(* IEC 61131-3 sources: Test-Git_ESME26/TestProgettoESME_26.fbsproj/PacDriveLib Migration/Motion/Homing/PDL_FB_Home.fb.st^, 21 files *)

(* ---- CallFb.meth.st ---- *)
{attribute 'conditionalshow_all_locals'}
METHOD PRIVATE CallFb
VAR_INPUT
END_VAR

CASE etHomeOpMode OF
	PDL_ET_HomeOpMode.TouchProbe:	(* HomeTP *)
		IF (stReducedVelocity_loc.i_xEnableReducedVelocity AND NOT stReducedVelocity_loc.i_xOnlyLimitCheck) THEN
			lrUsedVelocity := MIN(stReducedVelocity_loc.i_lrMaxReducedVelocity, stTouchProbe_loc.i_lrVel);
		ELSE
			lrUsedVelocity := stTouchProbe_loc.i_lrVel;
		END_IF
		fbHomeTP(	i_xEnable			:= xFbEnable,
					i_ifDrive			:= i_ifDrive,
					i_ifTouchProbe		:= stTouchProbe_loc.i_ifTouchProbe,
					i_etMode			:= etHomeTpMode,
					i_lrOffset			:= stTouchProbe_loc.i_lrOffset,
					i_lrMaxTravel		:= stTouchProbe_loc.i_lrMaxTravel,
					i_lrHomePosition	:= stTouchProbe_loc.i_lrHomePosition,
					i_lrVel				:= lrUsedVelocity,
					i_lrAcc				:= stTouchProbe_loc.i_lrAcc,
					i_lrDec				:= stTouchProbe_loc.i_lrDec,
					i_lrJerk			:= stTouchProbe_loc.i_lrJerk,
					i_xHwLimitNeg		:= i_xHwLimitNeg,
					i_xHwLimitPos		:= i_xHwLimitPos,
					i_xRotativeSystem	:= stTouchProbe_loc.i_xRotativeSystem,
					i_xStart			:= TRUE,
					q_xActive			=> xFbActive,
					q_xReady			=> ,
					q_etDiag			=> THIS^.etDiagBuffer,
					q_etDiagExt			=> ,
					q_sMsg				=> ,
					q_xMotionInstructionActive => ,
					q_lrPosition		=> ,
					q_xHomeOk			=> xFbHomeOk);
		THIS^.HomeTpDiagTranslation();

	PDL_ET_HomeOpMode.Sensor:	(* HomeIN *)
		IF (stReducedVelocity_loc.i_xEnableReducedVelocity AND NOT stReducedVelocity_loc.i_xOnlyLimitCheck) THEN
			lrUsedVelocity := MIN(stReducedVelocity_loc.i_lrMaxReducedVelocity, stSensor_loc.i_lrVel);
		ELSE
			lrUsedVelocity := stSensor_loc.i_lrVel;
		END_IF
		THIS^.fbHomeIn(	i_xEnable			:= xFbEnable,
					i_ifDrive			:= i_ifDrive,
					i_xSensor			:= stSensor_loc.i_xSensor,
					i_etMode			:= etHomeInMode,
					i_lrOffset			:= stSensor_loc.i_lrOffset,
					i_lrMaxTravel		:= stSensor_loc.i_lrMaxTravel,
					i_lrHomePosition	:= stSensor_loc.i_lrHomePosition,
					i_lrVel				:= lrUsedVelocity,
					i_lrAcc				:= stSensor_loc.i_lrAcc,
					i_lrDec				:= stSensor_loc.i_lrDec,
					i_lrJerk			:= stSensor_loc.i_lrJerk,
					i_xHwLimitNeg		:= i_xHwLimitNeg,
					i_xHwLimitPos		:= i_xHwLimitPos,
					i_xRotativeSystem	:= stSensor_loc.i_xRotativeSystem,
					i_xStart			:= xStartHomeIn,
					q_xActive			=> xFbActive,
					q_xReady			=> ,
					q_etDiag			=> THIS^.etDiagBuffer,
					q_etDiagExt			=> ,
					q_sMsg				=> ,
					q_xMotionInstructionActive => ,
					q_lrPosition		=> ,
					q_xHomeOk			=> xFbHomeOk);
		THIS^.HomeInDiagTranslation();

	PDL_ET_HomeOpMode.LimitSwitch:	(* HomeLS *)
		IF (stReducedVelocity_loc.i_xEnableReducedVelocity AND NOT stReducedVelocity_loc.i_xOnlyLimitCheck) THEN
			lrUsedVelocity := MIN(stReducedVelocity_loc.i_lrMaxReducedVelocity, stLimitSwitch_loc.i_lrVel);
		ELSE
			lrUsedVelocity := stLimitSwitch_loc.i_lrVel;
		END_IF
		IF (stLimitSwitch_loc.i_lrLowVel = 0.0) THEN
			lrLowVelocity := lrUsedVelocity;
		ELSE
			IF (stReducedVelocity_loc.i_xEnableReducedVelocity AND NOT stReducedVelocity_loc.i_xOnlyLimitCheck) THEN
				lrLowVelocity := MIN(stReducedVelocity_loc.i_lrMaxReducedVelocity, stLimitSwitch_loc.i_lrLowVel);
			ELSE
				lrLowVelocity := stLimitSwitch_loc.i_lrLowVel;
			END_IF
		END_IF
		fbHomeLS(	i_xEnable			:= xFbEnable,
					i_ifDrive			:= i_ifDrive,
					i_etMode			:= etHomeLimitSwitchMode,
					i_lrOffset			:= stLimitSwitch_loc.i_lrOffset,
					i_lrMaxTravel		:= stLimitSwitch_loc.i_lrMaxTravel,
					i_lrHomePosition	:= stLimitSwitch_loc.i_lrHomePosition,
					i_lrVel				:= lrUsedVelocity,
					i_lrLowVel			:= lrLowVelocity,
					i_lrAcc				:= stLimitSwitch_loc.i_lrAcc,
					i_lrDec				:= stLimitSwitch_loc.i_lrDec,
					i_lrJerk			:= stLimitSwitch_loc.i_lrJerk,
					i_xHwLimitNeg		:= i_xHwLimitNeg,
					i_xHwLimitPos		:= i_xHwLimitPos,
					i_xStart			:= TRUE,
					q_xActive			=> xFbActive,
					q_xReady			=> ,
					q_etDiag			=> THIS^.etDiagBuffer,
					q_etDiagExt			=> ,
					q_sMsg				=> ,
					q_xMotionInstructionActive => ,
					q_lrPosition		=> ,
					q_xHomeOk			=> xFbHomeOk);
		THIS^.HomeLSDiagTranslation();

	PDL_ET_HomeOpMode.Torque:	(* HomeTorque *)
		IF (stReducedVelocity_loc.i_xEnableReducedVelocity AND NOT stReducedVelocity_loc.i_xOnlyLimitCheck) THEN
			lrUsedVelocity := MIN(stReducedVelocity_loc.i_lrMaxReducedVelocity, stTorque_loc.i_lrVel);
		ELSE
			lrUsedVelocity := stTorque_loc.i_lrVel;
		END_IF
		fbHomeTorque(	i_xEnable			:= xFbEnable,
						i_ifDrive			:= i_ifDrive,
						i_lrMaxTorque		:= stTorque_loc.i_lrMaxTorque,
						i_diTorqueTime		:= stTorque_loc.i_diTorqueTime,
						i_lrLowLimit		:= -2147483648.0,
						i_lrHighLimit		:= 2147483648.0,
						i_etMode			:= etHomeTorqueMode,
						i_lrOffset			:= stTorque_loc.i_lrOffset,
						i_lrMaxTravel		:= stTorque_loc.i_lrMaxTravel,
						i_lrHomePosition	:= stTorque_loc.i_lrHomePosition,
						i_lrVel				:= lrUsedVelocity,
						i_lrAcc				:= stTorque_loc.i_lrAcc,
						i_lrDec				:= stTorque_loc.i_lrDec,
						i_lrJerk			:= stTorque_loc.i_lrJerk,
						i_xStart			:= TRUE,
						q_xActive			=> xFbActive,
						q_xReady			=> ,
						q_etDiag			=> THIS^.etDiagBuffer,
						q_etDiagExt			=> ,
						q_sMsg				=> ,
						q_xMotionInstructionActive => ,
						q_lrPosition		=> ,
						q_xHomeOk			=> xFbHomeOk);
		THIS^.HomeTorqueDiagTranslation();

	PDL_ET_HomeOpMode.Force:	(* HomeForce *)
			;

	PDL_ET_HomeOpMode.MoveOnPos:	(* Home to a Position *)
		IF (stReducedVelocity_loc.i_xEnableReducedVelocity AND NOT stReducedVelocity_loc.i_xOnlyLimitCheck) THEN
			lrUsedVelocity := MIN(stReducedVelocity_loc.i_lrMaxReducedVelocity, stMoveOnPos_loc.i_lrVel);
		ELSE
			lrUsedVelocity := stMoveOnPos_loc.i_lrVel;
		END_IF

		THIS^.fbVarioPosJerk(	i_xEnable			:= xFbEnable,
						i_ifDrive			:= i_ifDrive,
						i_xStart			:= fbVarioPosJerk.q_xActive AND TRUE,
						i_xStop				:= FALSE,
						i_lrTarget			:= lrPositionOpmMoveOnPos,
						i_lrVel				:= lrUsedVelocity,
						i_lrAcc				:= stMoveOnPos_loc.i_lrAcc,
						i_lrDec				:= stMoveOnPos_loc.i_lrDec,
						i_lrJerk			:= stMoveOnPos_loc.i_lrJerk,
						i_etPosMode			:= SEL(stMoveOnPos_loc.i_xRotativeSystem, PDL_ET_PosMode.Absolute, PDL_ET_PosMode.Relative),
						q_xActive			=> xFbActive,
						q_xReady			=> ,
						q_etDiag			=> THIS^.etDiagBuffer,
						q_etDiagExt			=> ,
						q_sMsg				=> ,
						q_xMotionInstructionActive => ,
						q_lrPosition		=> ,
						q_xInPosition		=> xFbHomeOk);

		THIS^.HomeMoveOnPosDiagTranslation();

		fbTrigStop(CLK:= xFbEnable AND (i_ifDrive.etAxisState = MOIN.ET_AxisState.Stopping));
		IF fbTrigStop.Q THEN
			xControllerStop :=  TRUE;
			xFbEnable := FALSE;
		END_IF

		// Clean up as soon as VarioPos is finished
		IF NOT xFbActive THEN
			// check, if VarioPos was aborted by MC_Stop OR MC_Halt
			IF xControllerStop THEN
				SetDiagOutput(	i_etDiag	:= GD.ET_Diag.HomingFailed,
								i_etDiagExt := PDL_ET_DiagExt.OutsideExecutionOfControllerStopSet,
								i_sMsg		:= 'MC_Stop OR MC_Halt was executed during homing active');
			ELSE
				IF stMoveOnPos_loc.i_lrPeriod > 0 AND stMoveOnPos_loc.i_xRotativeSystem THEN
					THIS^.fbSetPosIntern(
						Axis     := i_ifDrive,
						Position := stMoveOnPos_loc.i_lrTarget,
						Relative := FALSE,
						Execute  := TRUE);

					IF THIS^.fbSetPosIntern.Error THEN
							SetDiagOutput(	i_etDiag	:= GD.ET_Diag.UnexpectedProgramBehavior,
											i_etDiagExt := PDL_ET_DiagExt.UnexpectedFeedback,
											i_sMsg      := CONCAT('FB_Home error: MC_Setposition.ErrorID: ', PLCO.FC_EtResultToString(THIS^.fbSetPosIntern.ErrorID)));
					END_IF
					THIS^.fbSetPosIntern(Execute  := FALSE);
				END_IF
			END_IF
		END_IF

	PDL_ET_HomeOpMode.WritePos:	(* HomeAbs *)
		fbHomeAbs(	i_xEnable			:= xFbEnable,
					i_xExecute			:= TRUE,
					i_ifDrive			:= i_ifDrive,
					i_lrHomePosition	:= stWritePos_loc.i_lrHomePosition,
					i_lrAbsEncOffset	:= stWritePos_loc.i_lrAbsEncOffset,
					i_lrUserPeriod		:= stWritePos_loc.i_lrUserPeriod,
					q_xActive			=> xFbActive,
					q_xReady			=> ,
					q_xBusy				=> ,
					q_xDone				=> ,
					q_etDiag			=> THIS^.etDiagBuffer,
					q_etDiagExt			=> ,
					q_sMsg				=> ,
					q_xDisableDrive		=> q_xDisableDrive,
					q_lrPosition		=> ,
					q_xHomeOk			=> xFbHomeOk);
		THIS^.HomeWritePosDiagTranslation();

	PDL_ET_HomeOpMode.SetPos:	(* HomeSetPos *)
		THIS^.fbSetpos(	i_xEnable				:= xFbEnable,
					i_xExecute				:= TRUE,
					i_ifDrive				:= i_ifDrive,
					i_etMode				:= etHomeSetPosMode,
					i_lrHomePosition		:= stSetPos_loc.i_lrHomePosition,
					i_lrEncoderPosition		:= stSetPos_loc.i_lrEncoderPosition,
					i_lrAbsEncOffset		:= stSetPos_loc.i_lrAbsEncOffset,
					i_lrUserPeriod			:= stSetPos_loc.i_lrUserPeriod,
					i_lrRestoreWindow		:= stSetPos_loc.i_lrRestoreWindow,
					i_pstRestorePosRetain	:= stSetPos_loc.iq_pstRestorePosRetain,
					iq_lencEncoder			:= stSetPos_loc.iq_lencAxis,
					q_xActive				=> xFbActive,
					q_xReady				=> ,
					q_xBusy					=> ,
					q_xDone					=> ,
					q_etDiag				=> THIS^.etDiagBuffer,
					q_etDiagExt				=> ,
					q_sMsg					=> ,
					q_lrPosition			=> ,
					q_lrEncoderPosition		=> ,
					q_xHomeOk				=> xFbHomeOk);
		THIS^.HomeSetPosDiagTranslation();
END_CASE
IF NOT xFbActive THEN
	THIS^.etHomeOpMode := PDL_ET_HomeOpMode.NoOp;
END_IF

(* ---- DriveAndLencCheck.meth.st ---- *)
METHOD Private DriveAndLencCheck : BOOL
VAR_INPUT
END_VAR

//Check if used Axis and/or Logical Encoder are valid Elements of PLC-Configuration
		//Mode with Axis
	IF		THIS^.i_etMode = PDL_ET_HomeMode.PosDirectionPosEdgeTp
		OR	THIS^.i_etMode = PDL_ET_HomeMode.NegDirectionPosEdgeTp
		OR	THIS^.i_etMode = PDL_ET_HomeMode.NegDirectionNegEdgeTp
		OR	THIS^.i_etMode = PDL_ET_HomeMode.PosDirectionNegEdgeTp
		OR	THIS^.i_etMode = PDL_ET_HomeMode.PosDirectionPosEdgeSensor
		OR	THIS^.i_etMode = PDL_ET_HomeMode.NegDirectionPosEdgeSensor
		OR	THIS^.i_etMode = PDL_ET_HomeMode.NegDirectionNegEdgeSensor
		OR	THIS^.i_etMode = PDL_ET_HomeMode.PosDirectionNegEdgeSensor
		OR	THIS^.i_etMode = PDL_ET_HomeMode.PosDirectionPosEdgeHWLimitPos
		OR	THIS^.i_etMode = PDL_ET_HomeMode.NegDirectionPosEdgeHWLimitNeg
		OR	THIS^.i_etMode = PDL_ET_HomeMode.NegDirectionNegEdgeHWLimitNeg
		OR	THIS^.i_etMode = PDL_ET_HomeMode.PosDirectionNegEdgeHWLimitPos
		OR	THIS^.i_etMode = PDL_ET_HomeMode.PosDirectionMaxTorque
		OR	THIS^.i_etMode = PDL_ET_HomeMode.NegDirectionMaxTorque
		OR	THIS^.i_etMode = PDL_ET_HomeMode.MoveOnPosAbs
		OR	THIS^.i_etMode = PDL_ET_HomeMode.SetPosAxisPosition
		OR	THIS^.i_etMode = PDL_ET_HomeMode.RestorePosFromAxisEncoder
		OR	THIS^.i_etMode = PDL_ET_HomeMode.RestorePosFromRetain
		OR	THIS^.i_etMode = PDL_ET_HomeMode.WriteAxisEncoder THEN

			IF i_ifDrive = 0 THEN
					SetDiagOutput(	i_etDiag	:= GD.ET_Diag.InputParameterInvalid,
									i_etDiagExt := PDL_ET_DiagExt.DriveInvalid,
									i_sMsg		:= 'i_ifDrive = 0');
			END_IF

				//Mode with Lenc
	ELSIF THIS^.i_etMode = PDL_ET_HomeMode.SetPosLogEncoderPosition THEN
			IF THIS^.stSetPos_loc.iq_lencAxis = 0 THEN
				SetDiagOutput(	i_etDiag	:= GD.ET_Diag.InputParameterInvalid,
								i_etDiagExt := PDL_ET_DiagExt.LencInvalid,
								i_sMsg		:= 'iq_lencAxis = 0');
			END_IF

		//Mode with Axis and Lenc
	ELSIF THIS^.i_etMode = PDL_ET_HomeMode.SetPosAxisAndLogEncoderPosition THEN
			IF i_ifDrive = 0 THEN
					SetDiagOutput(	i_etDiag	:= GD.ET_Diag.InputParameterInvalid,
									i_etDiagExt := PDL_ET_DiagExt.DriveInvalid,
									i_sMsg		:= 'i_ifDrive = 0');

			ELSIF THIS^.stSetPos_loc.iq_lencAxis = 0 THEN
				SetDiagOutput(	i_etDiag	:= GD.ET_Diag.InputParameterInvalid,
								i_etDiagExt := PDL_ET_DiagExt.LencInvalid,
								i_sMsg		:= 'iq_lencAxis = 0');
			END_IF
	END_IF

(* ---- HomeForceDiagTranslation.meth.st ---- *)
METHOD PRIVATE HomeForceDiagTranslation : BOOL
VAR
END_VAR

IF THIS^.xFbEnable AND THIS^.fbHomeForce.q_etDiag <> GD.ET_Diag.Ok THEN

	CASE THIS^.fbHomeForce.q_etDiagExt OF

		PDL_ET_DiagExt.ControllerInvalid,
		PDL_ET_DiagExt.DriveNotReady,
		PDL_ET_DiagExt.MaxForceNotFound,
		PDL_ET_DiagExt.AccRange,
		PDL_ET_DiagExt.DecRange,
		PDL_ET_DiagExt.DriveInvalid,
		PDL_ET_DiagExt.JerkRange,
		PDL_ET_DiagExt.MaxForceRange,
		PDL_ET_DiagExt.MaxTravelRange,
		PDL_ET_DiagExt.VelRange,
		PDL_ET_DiagExt.SercosNotInPhaseFour,
		PDL_ET_DiagExt.UnexpectedFeedback,
		PDL_ET_DiagExt.UnknownState:

			THIS^.sTempMsg 	:= SE_CTBX.FC_MultiConcat(  i_sString1 := 'Mode HomeForce: ',
												i_sString2 := THIS^.fbHomeForce.q_sMsg,
												i_sString3 := '',
												i_sString4 := '');
			SetDiagOutput(	i_etDiag	:= THIS^.fbHomeForce.q_etDiag,
							i_etDiagExt := THIS^.fbHomeForce.q_etDiagExt,
							i_sMsg		:= THIS^.sTempMsg);
	ELSE
		sTempMsg 	:= SE_CTBX.FC_MultiConcat(  i_sString1 := 'Mode HomeForce, PDL_FB_HomeForce: ' ,
										i_sString2 := PDL_FC_EtDiagExtToString(i_etDiagExt := THIS^.fbHomeForce.q_etDiagExt),
										i_sString3 := THIS^.fbHomeForce.q_sMsg,
										i_sString4 := '');
		SetDiagOutput(	i_etDiag	:= GD.ET_Diag.UnexpectedProgramBehavior,
						i_etDiagExt := PDL_ET_DiagExt.UnexpectedFeedback,
						i_sMsg		:= THIS^.sTempMsg);
	END_CASE

END_IF

(* ---- HomeInDiagTranslation.meth.st ---- *)
METHOD Private HomeInDiagTranslation : BOOL
VAR
END_VAR

IF THIS^.xFbEnable AND THIS^.fbHomeIn.q_etDiag <> GD.ET_Diag.Ok THEN

	CASE THIS^.fbHomeIn.q_etDiagExt OF
		PDL_ET_DiagExt.DriveNotReady,
		PDL_ET_DiagExt.SensorNotFound,
		PDL_ET_DiagExt.AccRange,
		PDL_ET_DiagExt.DecRange,
		PDL_ET_DiagExt.DriveInvalid,
		PDL_ET_DiagExt.JerkRange,
		PDL_ET_DiagExt.MaxTravelRange,
		PDL_ET_DiagExt.VelRange,
		PDL_ET_DiagExt.HwLimitNegReached,
		PDL_ET_DiagExt.HwLimitPosReached,
		PDL_ET_DiagExt.HwLimitNegStillActive,
		PDL_ET_DiagExt.HwLimitPosStillActive,
		PDL_ET_DiagExt.SercosNotInPhaseFour,
		PDL_ET_DiagExt.UnexpectedFeedback,
		PDL_ET_DiagExt.UnknownState:

			THIS^.sTempMsg 	:= SE_CTBX.FC_MultiConcat(  i_sString1 := 'Mode HomeIn: ',
												i_sString2 := THIS^.fbHomeIn.q_sMsg,
												i_sString3 := '',
												i_sString4 := '');
			SetDiagOutput(	i_etDiag	:= THIS^.fbHomeIn.q_etDiag,
							i_etDiagExt := THIS^.fbHomeIn.q_etDiagExt,
							i_sMsg		:= THIS^.sTempMsg);
	ELSE
		sTempMsg 	:= SE_CTBX.FC_MultiConcat(  i_sString1 := 'Mode HomeIn, PDL_FB_HomeIn: ' ,
										i_sString2 := PDL_FC_EtDiagExtToString(i_etDiagExt := THIS^.fbHomeIn.q_etDiagExt),
										i_sString3 := THIS^.fbHomeIn.q_sMsg,
										i_sString4 := '');
		SetDiagOutput(	i_etDiag	:= GD.ET_Diag.UnexpectedProgramBehavior,
						i_etDiagExt := PDL_ET_DiagExt.UnexpectedFeedback,
						i_sMsg		:= THIS^.sTempMsg);
	END_CASE

END_IF

(* ---- HomeLSDiagTranslation.meth.st ---- *)
METHOD Private HomeLSDiagTranslation : BOOL
VAR
END_VAR

IF THIS^.xFbEnable AND THIS^.fbHomeLS.q_etDiag <> GD.ET_Diag.Ok THEN

	CASE THIS^.fbHomeLS.q_etDiagExt OF

		PDL_ET_DiagExt.DriveNotReady,
		PDL_ET_DiagExt.SensorNotFound,
		PDL_ET_DiagExt.AccRange,
		PDL_ET_DiagExt.DecRange,
		PDL_ET_DiagExt.DriveInvalid,
		PDL_ET_DiagExt.JerkRange,
		PDL_ET_DiagExt.LowVelRange,
		PDL_ET_DiagExt.MaxTravelRange,
		PDL_ET_DiagExt.VelRange,
		PDL_ET_DiagExt.HwLimitNegReached,
		PDL_ET_DiagExt.HwLimitPosReached,
		PDL_ET_DiagExt.SercosNotInPhaseFour,
		PDL_ET_DiagExt.UnexpectedFeedback,
		PDL_ET_DiagExt.UnknownState:

			THIS^.sTempMsg 	:= SE_CTBX.FC_MultiConcat(  i_sString1 := 'Mode HomeLS: ',
														i_sString2 := THIS^.fbHomeLS.q_sMsg,
														i_sString3 := '',
														i_sString4 := '');
			SetDiagOutput(	i_etDiag	:= THIS^.fbHomeLS.q_etDiag,
							i_etDiagExt := THIS^.fbHomeLS.q_etDiagExt,
							i_sMsg		:= THIS^.sTempMsg);
	ELSE
		sTempMsg 	:= SE_CTBX.FC_MultiConcat(  i_sString1 := 'Mode HomeLS, PDL_FB_HomeLimitSwitch: ' ,
												i_sString2 := PDL_FC_EtDiagExtToString(i_etDiagExt := THIS^.fbHomeLS.q_etDiagExt),
												i_sString3 := THIS^.fbHomeLS.q_sMsg,
												i_sString4 := '');
		SetDiagOutput(	i_etDiag	:= GD.ET_Diag.UnexpectedProgramBehavior,
						i_etDiagExt := PDL_ET_DiagExt.UnexpectedFeedback,
						i_sMsg		:= THIS^.sTempMsg);
	END_CASE

END_IF

(* ---- HomeMoveOnPosDiagTranslation.meth.st ---- *)
METHOD PRIVATE HomeMoveOnPosDiagTranslation : BOOL
VAR
END_VAR

IF THIS^.xFbEnable AND THIS^.fbVarioPosJerk.q_etDiag <> GD.ET_Diag.Ok THEN

	CASE THIS^.fbVarioPosJerk.q_etDiagExt OF
		PDL_ET_DiagExt.DriveNotReady,
		PDL_ET_DiagExt.AccRange,
		PDL_ET_DiagExt.DecRange,
		PDL_ET_DiagExt.DriveInvalid,
		PDL_ET_DiagExt.JerkRange,
		PDL_ET_DiagExt.VelRange,
		PDL_ET_DiagExt.SercosNotInPhaseFour,
		PDL_ET_DiagExt.UnexpectedFeedback,
		PDL_ET_DiagExt.UnknownState:

			THIS^.sTempMsg 	:= SE_CTBX.FC_MultiConcat(  i_sString1 := 'Mode HomeMoveOnPos: ',
												i_sString2 := THIS^.fbVarioPosJerk.q_sMsg,
												i_sString3 := '',
												i_sString4 := '');
			SetDiagOutput(	i_etDiag	:= THIS^.fbVarioPosJerk.q_etDiag,
							i_etDiagExt := THIS^.fbVarioPosJerk.q_etDiagExt,
							i_sMsg		:= THIS^.sTempMsg);
	ELSE
		sTempMsg 	:= SE_CTBX.FC_MultiConcat(  i_sString1 := 'Mode HomeMoveOnPos, PDL_FB_VarioPosJerk: ' ,
										i_sString2 := PDL_FC_EtDiagExtToString(i_etDiagExt := THIS^.fbVarioPosJerk.q_etDiagExt),
										i_sString3 := THIS^.fbVarioPosJerk.q_sMsg,
										i_sString4 := '');
		SetDiagOutput(	i_etDiag	:= GD.ET_Diag.UnexpectedProgramBehavior,
						i_etDiagExt := PDL_ET_DiagExt.UnexpectedFeedback,
						i_sMsg		:= THIS^.sTempMsg);
	END_CASE

END_IF

(* ---- HomeSetPosDiagTranslation.meth.st ---- *)
METHOD Private HomeSetPosDiagTranslation : BOOL
VAR
END_VAR

IF THIS^.xFbEnable AND THIS^.fbSetpos.q_etDiag <> GD.ET_Diag.Ok THEN

	CASE THIS^.fbSetpos.q_etDiagExt OF
		PDL_ET_DiagExt.DriveEncoderInvalid,
		PDL_ET_DiagExt.RestoreInterrupted,
		PDL_ET_DiagExt.SercosNotInPhaseFour,
		PDL_ET_DiagExt.AbsEncOffsetRange,
		PDL_ET_DiagExt.CheckSumInvalid,
		PDL_ET_DiagExt.DataNVRamInvalid,
		PDL_ET_DiagExt.DriveInvalid,
		PDL_ET_DiagExt.LencInvalid,
		PDL_ET_DiagExt.PointerRestorePosRetainInvalid,
		PDL_ET_DiagExt.UserPeriodRange,
		PDL_ET_DiagExt.OutOfRestoreWindow,
		PDL_ET_DiagExt.UnexpectedFeedback,
		PDL_ET_DiagExt.UnknownMode,
		PDL_ET_DiagExt.UnknownState:
			THIS^.sTempMsg 	:= SE_CTBX.FC_MultiConcat(  i_sString1 := 'Mode HomeSetPos: ',
														i_sString2 := THIS^.fbSetpos.q_sMsg,
														i_sString3 := '',
														i_sString4 := '');
			SetDiagOutput(	i_etDiag	:= THIS^.fbSetpos.q_etDiag,
							i_etDiagExt := THIS^.fbSetpos.q_etDiagExt,
							i_sMsg		:= THIS^.sTempMsg);
	ELSE
		sTempMsg 	:= SE_CTBX.FC_MultiConcat(  i_sString1 := 'Mode HomeSetPos, PDL_FB_HomeSetPos: ' ,
												i_sString2 := PDL_FC_EtDiagExtToString(i_etDiagExt := THIS^.fbSetpos.q_etDiagExt),
												i_sString3 := THIS^.fbSetpos.q_sMsg,
												i_sString4 := '');
		SetDiagOutput(	i_etDiag	:= GD.ET_Diag.UnexpectedProgramBehavior,
						i_etDiagExt := PDL_ET_DiagExt.UnexpectedFeedback,
						i_sMsg		:= THIS^.sTempMsg);
	END_CASE

END_IF

(* ---- HomeTorqueDiagTranslation.meth.st ---- *)
METHOD PRIVATE HomeTorqueDiagTranslation : BOOL
VAR
END_VAR

IF THIS^.xFbEnable AND THIS^.fbHomeTorque.q_etDiag <> GD.ET_Diag.Ok THEN

	CASE THIS^.fbHomeTorque.q_etDiagExt OF

		PDL_ET_DiagExt.ControllerInvalid,
		PDL_ET_DiagExt.DriveNotReady,
		PDL_ET_DiagExt.MaxTorqueNotFound,
		PDL_ET_DiagExt.AccRange,
		PDL_ET_DiagExt.DecRange,
		PDL_ET_DiagExt.DriveInvalid,
		PDL_ET_DiagExt.JerkRange,
		PDL_ET_DiagExt.MaxTorqueRange,
		PDL_ET_DiagExt.MaxTravelRange,
		PDL_ET_DiagExt.VelRange,
		PDL_ET_DiagExt.SercosNotInPhaseFour,
		PDL_ET_DiagExt.UnexpectedFeedback,
		PDL_ET_DiagExt.UnknownState:

			THIS^.sTempMsg 	:= SE_CTBX.FC_MultiConcat(  i_sString1 := 'Mode HomeTorque: ',
												i_sString2 := THIS^.fbHomeTorque.q_sMsg,
												i_sString3 := '',
												i_sString4 := '');
			SetDiagOutput(	i_etDiag	:= THIS^.fbHomeTorque.q_etDiag,
							i_etDiagExt := THIS^.fbHomeTorque.q_etDiagExt,
							i_sMsg		:= THIS^.sTempMsg);
	ELSE
		sTempMsg 	:= SE_CTBX.FC_MultiConcat(  i_sString1 := 'Mode HomeTorque, PDL_FB_HomeTorque: ' ,
										i_sString2 := PDL_FC_EtDiagExtToString(i_etDiagExt := THIS^.fbHomeTorque.q_etDiagExt),
										i_sString3 := THIS^.fbHomeTorque.q_sMsg,
										i_sString4 := '');
		SetDiagOutput(	i_etDiag	:= GD.ET_Diag.UnexpectedProgramBehavior,
						i_etDiagExt := PDL_ET_DiagExt.UnexpectedFeedback,
						i_sMsg		:= THIS^.sTempMsg);
	END_CASE

END_IF

(* ---- HomeTpDiagTranslation.meth.st ---- *)
METHOD Private HomeTpDiagTranslation : BOOL
VAR
END_VAR

IF THIS^.xFbEnable AND THIS^.fbHomeTP.q_etDiag <> GD.ET_Diag.Ok THEN

	CASE THIS^.fbHomeTP.q_etDiagExt OF
		PDL_ET_DiagExt.DriveNotReady,
		PDL_ET_DiagExt.TouchProbeNotFound,
		PDL_ET_DiagExt.AccRange,
		PDL_ET_DiagExt.DecRange,
		PDL_ET_DiagExt.DriveInvalid,
		PDL_ET_DiagExt.JerkRange,
		PDL_ET_DiagExt.MaxTravelRange,
		PDL_ET_DiagExt.TouchProbeInvalid,
		PDL_ET_DiagExt.TouchProbeNotActive,
		PDL_ET_DiagExt.TouchProbeVirtual,
		PDL_ET_DiagExt.VelRange,
		PDL_ET_DiagExt.HwLimitNegReached,
		PDL_ET_DiagExt.HwLimitPosReached,
		PDL_ET_DiagExt.HwLimitNegStillActive,
		PDL_ET_DiagExt.HwLimitPosStillActive,
		PDL_ET_DiagExt.SercosNotInPhaseFour,
		PDL_ET_DiagExt.UnexpectedFeedback,
		PDL_ET_DiagExt.UnknownState :

			THIS^.sTempMsg 	:= SE_CTBX.FC_MultiConcat(  i_sString1 := 'Mode HomeTP: ',
														i_sString2 := THIS^.fbHomeTP.q_sMsg,
														i_sString3 := '',
														i_sString4 := '');
			SetDiagOutput(	i_etDiag	:= THIS^.fbHomeTP.q_etDiag,
							i_etDiagExt := THIS^.fbHomeTP.q_etDiagExt,
							i_sMsg		:= THIS^.sTempMsg);
	ELSE
		sTempMsg 	:= SE_CTBX.FC_MultiConcat(  i_sString1 := 'Mode HomeTP, PDL_FB_HomeTp: ' ,
												i_sString2 := PDL_FC_EtDiagExtToString(i_etDiagExt := THIS^.fbHomeTP.q_etDiagExt),
												i_sString3 := THIS^.fbHomeTP.q_sMsg,
												i_sString4 := '');
		SetDiagOutput(	i_etDiag	:= GD.ET_Diag.UnexpectedProgramBehavior,
						i_etDiagExt := PDL_ET_DiagExt.UnexpectedFeedback,
						i_sMsg		:= THIS^.sTempMsg);
	END_CASE

END_IF

(* ---- HomeWritePosDiagTranslation.meth.st ---- *)
METHOD Private HomeWritePosDiagTranslation : BOOL
VAR
END_VAR

IF THIS^.xFbEnable AND THIS^.fbHomeAbs.q_etDiag <> GD.ET_Diag.Ok THEN

	CASE THIS^.fbHomeAbs.q_etDiagExt OF

		PDL_ET_DiagExt.SercosInterfaceInvalid,
		PDL_ET_DiagExt.DriveEncoderInvalid,
		PDL_ET_DiagExt.DriveIsMoving,
		PDL_ET_DiagExt.DriveNotDisabled,
		PDL_ET_DiagExt.NoAccessToEEPROM,
		PDL_ET_DiagExt.ProgrammingInProgress,
		PDL_ET_DiagExt.ProgrammingInvalidEEPROM,
		PDL_ET_DiagExt.AbsEncOffsetRange,
		PDL_ET_DiagExt.DriveInvalid,
		PDL_ET_DiagExt.UserPeriodRange,
		PDL_ET_DiagExt.SercosNotInPhaseFour,
		PDL_ET_DiagExt.EncoderWriteTimeOut,
		PDL_ET_DiagExt.UnexpectedFeedback,
		PDL_ET_DiagExt.UnknownState:

			THIS^.sTempMsg 	:= SE_CTBX.FC_MultiConcat(  i_sString1 := 'Mode HomeWritePos: ',
												i_sString2 := THIS^.fbHomeAbs.q_sMsg,
												i_sString3 := '',
												i_sString4 := '');
			SetDiagOutput(	i_etDiag	:= THIS^.fbHomeAbs.q_etDiag,
							i_etDiagExt := THIS^.fbHomeAbs.q_etDiagExt,
							i_sMsg		:= THIS^.sTempMsg);
	ELSE
		sTempMsg 	:= SE_CTBX.FC_MultiConcat(  i_sString1 := 'Mode HomeWritePos, PDL_FB_HomeAbs: ' ,
										i_sString2 := PDL_FC_EtDiagExtToString(i_etDiagExt := THIS^.fbHomeAbs.q_etDiagExt),
										i_sString3 := THIS^.fbHomeAbs.q_sMsg,
										i_sString4 := '');
		SetDiagOutput(	i_etDiag	:= GD.ET_Diag.UnexpectedProgramBehavior,
						i_etDiagExt := PDL_ET_DiagExt.UnexpectedFeedback,
						i_sMsg		:= THIS^.sTempMsg);
	END_CASE

END_IF

(* ---- RegisterLoggerPoint.meth.st ---- *)
{attribute 'conditionalshow_all_locals'}
METHOD PUBLIC RegisterLoggerPoint
VAR_INPUT
	i_ifParent		: APL.IF_LoggerPoint;
	i_sName			: STRING[80];
END_VAR
VAR_OUTPUT
	q_etDiag		: GD.ET_Diag := GD.ET_Diag.Ok;
	q_etDiagExt		: PDL_ET_DiagExt := PDL_ET_DiagExt.Ok;
END_VAR
VAR
	etDiagBuffer		: GD.ET_Diag;
	etDiagExtBufferAPL	: APL.ET_DiagExt;
END_VAR

THIS^.fbLoggerPoint.RegisterLoggerPoint(	i_ifParent		:= i_ifParent,
											i_sName			:= i_sName,
											i_sType			:= 'FB_Home',
											i_sSource		:= 'PDL',
											q_etDiag		=> etDiagBuffer,
											q_etDiagExt		=> etDiagExtBufferAPL);
IF (etDiagBuffer <> GD.ET_Diag.Ok) THEN
	CASE etDiagExtBufferAPL OF
		APL.ET_DiagExt.ParentInvalid:
			q_etDiag := GD.ET_Diag.InputParameterInvalid;
			q_etDiagExt := PDL_ET_DiagExt.ParentInvalid;

		APL.ET_DiagExt.ParentNotRegistered:
			q_etDiag := GD.ET_Diag.InputParameterInvalid;
			q_etDiagExt := PDL_ET_DiagExt.ParentNotRegistered;

		APL.ET_DiagExt.MaxNumberOfLoggerPointsExeeded:
			q_etDiag := GD.ET_Diag.InputParameterInvalid;
			q_etDiagExt := PDL_ET_DiagExt.MaxNumberOfLoggerPointsExeeded;

	ELSE
		q_etDiag := GD.ET_Diag.UnexpectedProgramBehavior;
		q_etdiagExt := PDL_ET_DiagExt.UnexpectedDiagExt;
	END_CASE
END_IF

(* ---- SetDiagOutput.meth.st ---- *)
METHOD PRIVATE SetDiagOutput : BOOL
VAR_INPUT
	i_etDiag	: GD.ET_Diag;
	i_etDiagExt	: PDL_ET_DiagExt;
	i_sMsg		: STRING[80];
END_VAR
VAR
END_VAR

IF i_etDiag <> GD.ET_Diag.Ok THEN
	q_xReady := FALSE;
END_IF
IF q_etDiag = GD.ET_Diag.OK OR i_etDiagExt = PDL_ET_DiagExt.Disabled THEN
	q_etDiag := i_etDiag;
	q_etDiagExt := i_etDiagExt;
	q_sMsg := i_sMsg;

	IF(i_etDiag = GD.ET_Diag.Ok) AND (THIS^.fbLoggerPoint.etLogLevel >= APL.ET_LogLevel.StatusMessage) THEN
		THIS^.fbLoggerPoint.AddLogEntry(	i_etLogLevel	:= APL.ET_LogLevel.StatusMessage,
											i_etDiag		:= q_etDiag,
											i_udiDiagExt	:= q_etDiagExt,
											i_sMessage		:= SE_CTBX.FC_MultiConcat(	i_sString1	:= Standard.CONCAT('ET_Diag: ', GD.FC_EtDiagToString(q_etDiag)),
																				i_sString2	:= Standard.CONCAT(' ET_DiagExt: ', PDL_FC_EtDiagExtToString(q_etDiagExt)),
																				i_sString3	:= Standard.CONCAT(' sMsg: ', q_sMsg),
																				i_sString4	:= ''),
											q_etDiag		:= ,	// ignore result
											q_etDiagExt		:= );	// ignore result
	ELSIF(i_etDiag = GD.ET_Diag.UnexpectedProgramBehavior) AND (THIS^.fbLoggerPoint.etLogLevel >= APL.ET_LogLevel.CriticalException) THEN
		THIS^.fbLoggerPoint.AddLogEntry(	i_etLogLevel	:= APL.ET_LogLevel.CriticalException,
											i_etDiag		:= q_etDiag,
											i_udiDiagExt	:= q_etDiagExt,
											i_sMessage		:= SE_CTBX.FC_MultiConcat(	i_sString1	:= Standard.CONCAT('ET_Diag: ', GD.FC_EtDiagToString(q_etDiag)),
																				i_sString2	:= Standard.CONCAT(' ET_DiagExt: ', PDL_FC_EtDiagExtToString(q_etDiagExt)),
																				i_sString3	:= Standard.CONCAT(' sMsg: ', q_sMsg),
																				i_sString4	:= ''),
											q_etDiag		:= ,	// ignore result
											q_etDiagExt		:= );	// ignore result
	ELSIF(i_etDiag <> GD.ET_Diag.Ok) AND (THIS^.fbLoggerPoint.etLogLevel >= APL.ET_LogLevel.Exception) THEN
		THIS^.fbLoggerPoint.AddLogEntry(	i_etLogLevel	:= APL.ET_LogLevel.Exception,
											i_etDiag		:= q_etDiag,
											i_udiDiagExt	:= q_etDiagExt,
											i_sMessage		:= SE_CTBX.FC_MultiConcat(	i_sString1	:= Standard.CONCAT('ET_Diag: ', GD.FC_EtDiagToString(q_etDiag)),
																				i_sString2	:= Standard.CONCAT(' ET_DiagExt: ', PDL_FC_EtDiagExtToString(q_etDiagExt)),
																				i_sString3	:= Standard.CONCAT(' sMsg: ', q_sMsg),
																				i_sString4	:= ''),
											q_etDiag		:= ,	// ignore result
											q_etDiagExt		:= );	// ignore result
	END_IF
END_IF

IF q_etDiag <> GD.ET_Diag.OK THEN
	THIS^.xFbEnable	:= FALSE;
	THIS^.q_xReady := FALSE;
	THIS^.q_xHomeOK := FALSE;
	IF xEnableFlag THEN
		THIS^.etHomeState := PDL_ET_HomeState.ExceptionOrIdle;
	END_IF
END_IF

(* ---- stForce.prop.st ---- *)
PROPERTY stForce : PDL_ST_HomeForce
__GETTERDECLARATION__
VAR
END_VAR
__GETTERIMPLEMENTATION__
stForce:= THIS^.stForce_loc;
__SETTERDECLARATION__
VAR
END_VAR
__SETTERIMPLEMENTATION__
THIS^.stForce_loc := stForce;

(* ---- stLimitSwitch.prop.st ---- *)
PROPERTY stLimitSwitch : PDL_ST_HomeLimitSwitch
__SETTERDECLARATION__
VAR
END_VAR
__SETTERIMPLEMENTATION__
THIS^.stLimitSwitch_loc := stLimitSwitch;
__GETTERDECLARATION__
VAR
END_VAR
__GETTERIMPLEMENTATION__
stLimitSwitch := THIS^.stLimitSwitch_loc;

(* ---- stMoveOnPos.prop.st ---- *)
PROPERTY stMoveOnPos : PDL_ST_HomeMoveOnPos
__SETTERDECLARATION__
VAR
END_VAR
__SETTERIMPLEMENTATION__
THIS^.stMoveOnPos_loc := stMoveOnPos;
__GETTERDECLARATION__
VAR
END_VAR
__GETTERIMPLEMENTATION__
stMoveOnPos := THIS^.stMoveOnPos_loc;

(* ---- stReducedVelocity.prop.st ---- *)
PROPERTY stReducedVelocity : PDL_ST_ReducedVelocity
__SETTERDECLARATION__
VAR
END_VAR
__SETTERIMPLEMENTATION__
THIS^.stReducedVelocity_loc := stReducedVelocity;
__GETTERDECLARATION__
VAR
END_VAR
__GETTERIMPLEMENTATION__
stReducedVelocity := THIS^.stReducedVelocity_loc;

(* ---- stSensor.prop.st ---- *)
PROPERTY stSensor : PDL_ST_HomeIn
__SETTERDECLARATION__
VAR
END_VAR
__SETTERIMPLEMENTATION__
THIS^.stSensor_loc := stSensor;
__GETTERDECLARATION__
VAR
END_VAR
__GETTERIMPLEMENTATION__
stSensor := THIS^.stSensor_loc;

(* ---- stSetPos.prop.st ---- *)
PROPERTY stSetPos : PDL_ST_HomeSetPos
__SETTERDECLARATION__
VAR
END_VAR
__SETTERIMPLEMENTATION__
THIS^.stSetPos_loc := stSetPos;
__GETTERDECLARATION__
VAR
END_VAR
__GETTERIMPLEMENTATION__
stSetPos := THIS^.stSetPos_loc;

(* ---- stTorque.prop.st ---- *)
PROPERTY stTorque : PDL_ST_HomeTorque
__GETTERDECLARATION__
VAR
END_VAR
__GETTERIMPLEMENTATION__
stTorque := THIS^.stTorque_loc;
__SETTERDECLARATION__
VAR
END_VAR
__SETTERIMPLEMENTATION__
THIS^.stTorque_loc := stTorque;

(* ---- stTouchProbe.prop.st ---- *)
PROPERTY stTouchProbe : PDL_ST_HomeTp
__SETTERDECLARATION__
VAR
END_VAR
__SETTERIMPLEMENTATION__
THIS^.stTouchProbe_loc := stTouchProbe;
__GETTERDECLARATION__
VAR
END_VAR
__GETTERIMPLEMENTATION__
stTouchProbe := THIS^.stTouchProbe_loc;

(* ---- stWritePos.prop.st ---- *)
PROPERTY stWritePos : PDL_ST_HomeWritePos
__SETTERDECLARATION__
VAR
END_VAR
__SETTERIMPLEMENTATION__
THIS^.stWritePos_loc := stWritePos;
__GETTERDECLARATION__
VAR
END_VAR
__GETTERIMPLEMENTATION__
stWritePos := THIS^.stWritePos_loc;
